{attribute 'qualified_only'}
{attribute 'strict'}
{attribute 'to_string'}
TYPE E_Line_Source :
(
	eNone := 0,
	eClose,
	eTank_A,
	eTank_B,
	eTapWater,
	eFillWater,
	eCIP,
	eDrain
);
END_TYPE

(* stored: Version 1.1.0.1, ProductVersion 3.1.4024.12
   DUT E_Line_Source: Id {0297a55d-f777-4926-8502-b778eb411f36} *)
